TYPE "ST_PressDemoParCfg"
VERSION : 0.1
   STRUCT
      SchemaVersion : UInt := 1;
      Timeout : Time := T#0MS;
   END_STRUCT;

END_TYPE

